% RSLogix 500 project PROGRAM_6.RSS, saved by version 8.30.00.16 %
PROJECT "UNTITLED"    % processor: Bul.1763 MicroLogix 1100 Series B %

PROGRAM FILES
  LAD 2 "MAIN"  3 rungs
  LAD 3 "IO"  2 rungs
  LAD 4 "HOURMETER"  9 rungs

DATA FILES
  O0 OUTPUT  4 elements
  I1 INPUT  6 elements
  S2 STATUS  66 elements
  B3 BINARY  1 elements
  T4 TIMER  1 elements
  C5 COUNTER  1 elements
  R6 CONTROL  1 elements
  N7 INTEGER  4 elements
  F8 FLOAT  1 elements

LADDER 2 "MAIN"
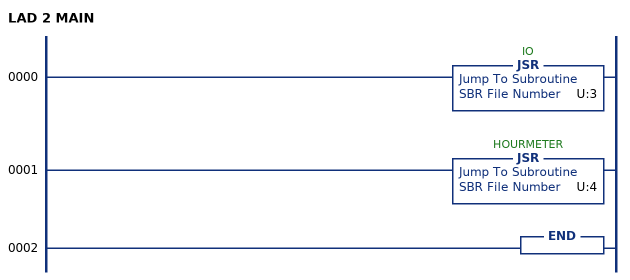
% Rung: 0 %
SOR JSR U:3 EOR
%   U:3  "IO" %
% Rung: 1 %
SOR JSR U:4 EOR
%   U:4  "HOURMETER" %
% Rung: 2 %
SOR END EOR

LADDER 3 "IO"
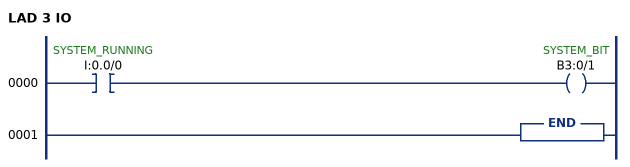
% Rung: 0 %
SOR XIC I:0.0/0 OTE B3:0/1 EOR
%   I:0.0/0  "SYSTEM_RUNNING" %
%   B3:0/1  "SYSTEM_BIT" %
% Rung: 1 %
SOR END EOR

LADDER 4 "HOURMETER"
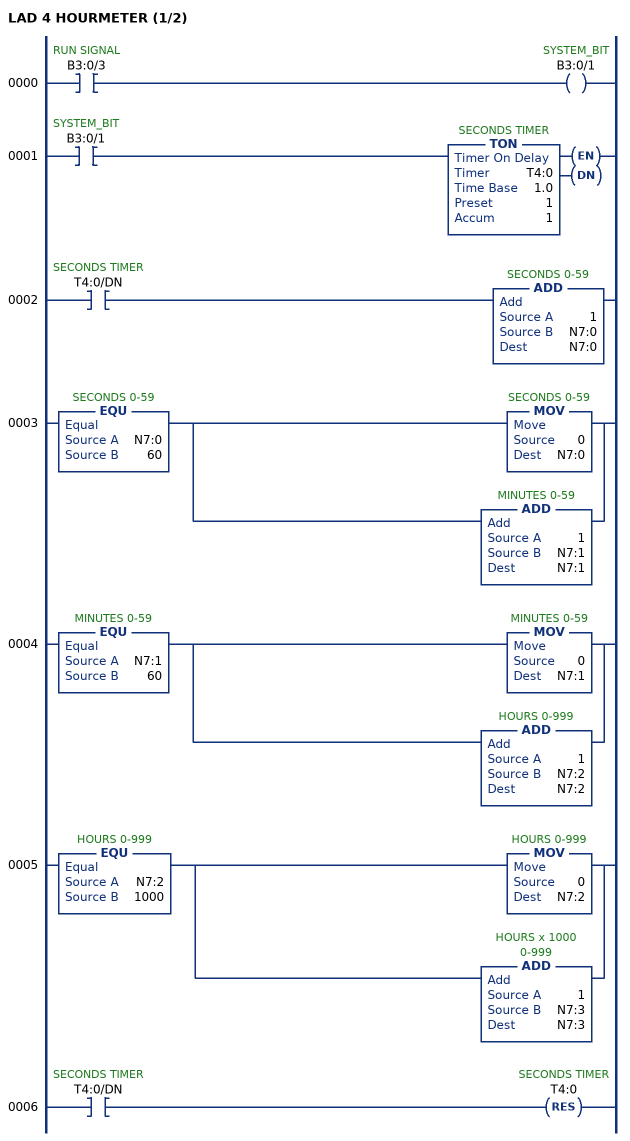
% Rung: 0 %
SOR XIC B3:0/3 OTE B3:0/1 EOR
%   B3:0/3  "RUN SIGNAL" %
%   B3:0/1  "SYSTEM_BIT" %
% Rung: 1 %
SOR XIC B3:0/1 TON T4:0 1.0 1 1 EOR
%   B3:0/1  "SYSTEM_BIT" %
%   T4:0  "SECONDS TIMER" %
% Rung: 2 %
SOR XIC T4:0/DN ADD 1 N7:0 N7:0 EOR
%   T4:0  "SECONDS TIMER" %
%   N7:0  "SECONDS 0-59" %
% Rung: 3 %
SOR EQU N7:0 60 BST MOV 0 N7:0 NXB ADD 1 N7:1 N7:1 BND EOR
%   N7:0  "SECONDS 0-59" %
%   N7:1  "MINUTES 0-59" %
% Rung: 4 %
SOR EQU N7:1 60 BST MOV 0 N7:1 NXB ADD 1 N7:2 N7:2 BND EOR
%   N7:1  "MINUTES 0-59" %
%   N7:2  "HOURS 0-999" %
% Rung: 5 %
SOR EQU N7:2 1000 BST MOV 0 N7:2 NXB ADD 1 N7:3 N7:3 BND EOR
%   N7:2  "HOURS 0-999" %
%   N7:3  "HOURS x 1000 0-999" %
% Rung: 6 %
SOR XIC T4:0/DN RES T4:0 EOR
%   T4:0  "SECONDS TIMER" %

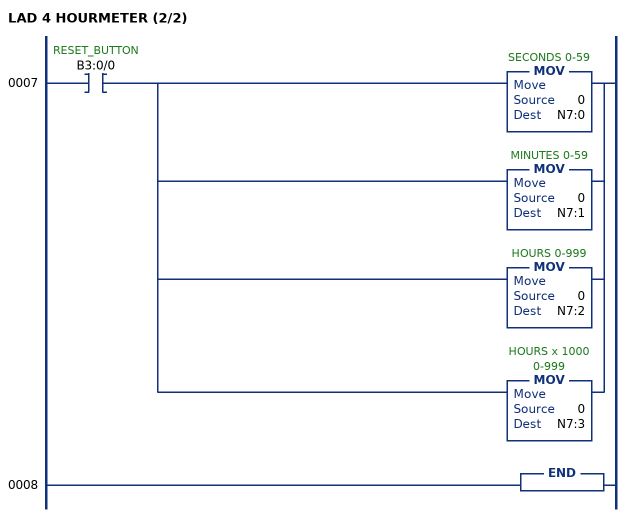
% Rung: 7 %
SOR XIC B3:0/0 BST MOV 0 N7:0 NXB MOV 0 N7:1 NXB MOV 0 N7:2 NXB MOV 0 N7:3 BND EOR
%   B3:0/0  RESET_BUTTON %
%   N7:0  "SECONDS 0-59" %
%   N7:1  "MINUTES 0-59" %
%   N7:2  "HOURS 0-999" %
%   N7:3  "HOURS x 1000 0-999" %
% Rung: 8 %
SOR END EOR

OTHER DOCUMENTED ADDRESSES
  C5:0  "SECONDS COUNTER"
  T4:0.ACC  "SECONDS ACC"
  T4:1  "MINUTES 0-59"

DATA TABLE (non-zero values as saved)
DATA B3
% B3:0 % 0X0002
DATA T4
% .PRE .ACC %
% T4:0 % 1 1
DATA N7
% N7:0 % 42 1 0 1
